(* IEC 61131-3 sources: SRCI_CLIENT_PLC/RobotLibrary/Library/Enumerations/Miscellaneous, 14 files *)

(* ---- AxisUnit.st ---- *)
{attribute 'qualified_only'}
{attribute 'to_string'}
{attribute 'strict'}
// -------------------------------------------------------------------------
//  SRCI Robot Library
// -------------------------------------------------------------------------
//
//  Object:      AxisUnit
//  Author:      Thorsten Brach
//  Date:        2025-03-23
//
//  Description:
//
//
//  Copyright:
//    (C) 2025 Thorsten Brach. All rights reserved
//             Licensed under the MIT License.
//
//  Disclaimer:
//    This project is provided without any guarantee and can be used for
//    private and commercial purposes. Any use is at the user’s
//    own risk and responsibility.
//
// -------------------------------------------------------------------------
TYPE AxisUnit :
(
  /// Axis unit is in degree [°]
	DEG := 0,
  /// Axis unit is in milli meter [mm]
	MM  := 1
)USINT;
END_TYPE

(* ---- CircPlane.st ---- *)
{attribute 'qualified_only'}
{attribute 'to_string'}
{attribute 'strict'}
// -------------------------------------------------------------------------
//  SRCI Robot Library
// -------------------------------------------------------------------------
//
//  Object:      CircPlane
//  Author:      Thorsten Brach
//  Date:        2024-06-01
//
//  Description:
//
//
//  Copyright:
//    (C) 2024 Thorsten Brach. All rights reserved
//             Licensed under the MIT License.
//
//  Disclaimer:
//    This project is provided without any guarantee and can be used for
//    private and commercial purposes. Any use is at the user’s
//    own risk and responsibility.
//
// -------------------------------------------------------------------------
TYPE CircPlane :
(
  /// x-z-plane
  XZ_PLANE := 0,
  /// y-z-plane
  YZ_PLANE := 1,
  /// x-y-plane
  XY_PLANE := 2
)SINT;
END_TYPE

(* ---- ComDirection.st ---- *)
{attribute 'qualified_only'}
{attribute 'to_string'}
{attribute 'strict'}
// -------------------------------------------------------------------------
//  SRCI Robot Library
// -------------------------------------------------------------------------
//
//  Object:      ComDirection
//  Author:      Thorsten Brach
//  Date:        2025-03-23
//
//  Description:
//
//
//  Copyright:
//    (C) 2025 Thorsten Brach. All rights reserved
//             Licensed under the MIT License.
//
//  Disclaimer:
//    This project is provided without any guarantee and can be used for
//    private and commercial purposes. Any use is at the user’s
//    own risk and responsibility.
//
// -------------------------------------------------------------------------
TYPE ComDirection :
(
  // communication direction PLC to Robot
	PLC_TO_ROB := 0,
  // communication direction Robot to PLC
	ROB_TO_PLC := 1
);
END_TYPE

(* ---- ControlHalfByte.st ---- *)
{attribute 'qualified_only'}
{attribute 'to_string'}
// -------------------------------------------------------------------------
//  SRCI Robot Library
// -------------------------------------------------------------------------
//
//  Object:      ControlHalfByte
//  Author:      Thorsten Brach
//  Date:        2024-06-01
//
//  Description:
//
//
//  Copyright:
//    (C) 2024 Thorsten Brach. All rights reserved
//             Licensed under the MIT License.
//
//  Disclaimer:
//    This project is provided without any guarantee and can be used for
//    private and commercial purposes. Any use is at the user’s
//    own risk and responsibility.
//
// -------------------------------------------------------------------------
TYPE ControlHalfByte :
(
  /// Default value, no control active
  NONE := 0,
  /// Initialization is requested by the client
  INITIALIZE := 1,
  /// Resume of operation is requested by the client
  RESUME := 2,
  /// Resetting of the RC is requested by the client. The RC must stop the motion, and clear all state.
  RESET := 3,
  /// Acknowledgement of a telegram state error
  ACK_ERROR := 4,
  /// Signaling that a client error occurred. The Server must respond by setting its RI state to NOT_INITIALIZED
  CLIENT_ERROR := 5
)BYTE;
END_TYPE

(* ---- ErrorReaction.st ---- *)
{attribute 'qualified_only'}
{attribute 'to_string'}
// -------------------------------------------------------------------------
//  SRCI Robot Library
// -------------------------------------------------------------------------
//
//  Object:      ErrorReaction
//  Author:      Thorsten Brach
//  Date:        2024-06-01
//
//  Description:
//
//
//  Copyright:
//    (C) 2024 Thorsten Brach. All rights reserved
//             Licensed under the MIT License.
//
//  Disclaimer:
//    This project is provided without any guarantee and can be used for
//    private and commercial purposes. Any use is at the user’s
//    own risk and responsibility.
//
// -------------------------------------------------------------------------
TYPE ErrorReaction :
(
  /// Abort and move Abort active move command and delete commands buffered in sequence Move robot by specified ErrorVector
  ABORT_AND_MOVE := 0,
  /// 1: Abort
  /// Abort active move command and delete commands buffered in sequence
  /// No additional movements
  ABORT := 1,
  /// 2: No reaction
  /// Error event is ignored by active move command
  NO_REACTION := 2
)USINT;
END_TYPE

(* ---- LoadMeasurementSteps.st ---- *)
{attribute 'qualified_only'}
{attribute 'to_string'}
// -------------------------------------------------------------------------
//  SRCI Robot Library
// -------------------------------------------------------------------------
//
//  Object:      LoadMeasurementSteps
//  Author:      Thorsten Brach
//  Date:        2024-06-01
//
//  Description:
//
//
//  Copyright:
//    (C) 2024 Thorsten Brach. All rights reserved
//             Licensed under the MIT License.
//
//  Disclaimer:
//    This project is provided without any guarantee and can be used for
//    private and commercial purposes. Any use is at the user’s
//    own risk and responsibility.
//
// -------------------------------------------------------------------------
TYPE LoadMeasurementSteps :
(
  /// • 0: Reset (default)
  /// Delete all positions saved on the RC
  RESET := 0,
  /// • 1: First position
  /// Save the first position for the load estimation with the required data
  FIRST_POSITION := 1,
  /// • 2: Second position
  /// Save the second position for the load estimation with the required data
  SECOND_POSITION := 2,
  /// • 3: Third position
  /// Save the third position for the load estimation with the required data
  THIRD_POSITION := 3,
  /// • 4: Fourth position
  /// Save the fourth position for the load estimation with the required data
  FOURTH_POSITION := 4,
  /// • 99: Load calculation
  /// Start the load calculation with the data saved in the four positions
  LOAD_CALCULATION := 99
)USINT;
END_TYPE

(* ---- PathChoice.st ---- *)
{attribute 'qualified_only'}
{attribute 'to_string'}
// -------------------------------------------------------------------------
//  SRCI Robot Library
// -------------------------------------------------------------------------
//
//  Object:      PathChoice
//  Author:      Thorsten Brach
//  Date:        2024-06-01
//
//  Description:
//
//
//  Copyright:
//    (C) 2024 Thorsten Brach. All rights reserved
//             Licensed under the MIT License.
//
//  Disclaimer:
//    This project is provided without any guarantee and can be used for
//    private and commercial purposes. Any use is at the user’s
//    own risk and responsibility.
//
// -------------------------------------------------------------------------
TYPE PathChoice :
(
  /// Clockwise movement of the circular path
  CLOCKWISE := 0,
  /// Counterclockwise movement of the circular path
  COUNTERCLOCKWISE := 1
)BYTE;
END_TYPE

(* ---- ReferenceElement.st ---- *)
{attribute 'qualified_only'}
{attribute 'to_string'}
// -------------------------------------------------------------------------
//  SRCI Robot Library
// -------------------------------------------------------------------------
//
//  Object:      ReferenceElement
//  Author:      Thorsten Brach
//  Date:        2024-06-01
//
//  Description:
//
//
//  Copyright:
//    (C) 2024 Thorsten Brach. All rights reserved
//             Licensed under the MIT License.
//
//  Disclaimer:
//    This project is provided without any guarantee and can be used for
//    private and commercial purposes. Any use is at the user’s
//    own risk and responsibility.
//
// -------------------------------------------------------------------------
TYPE ReferenceElement :
(
  /// 0 (default): Not used
  NOT_USED := 0,
  /// 1: X-Axis
  X_AXIS := 1,
  /// 2: Y-Axis
  Y_AXIS := 2,
  /// 3: Z-Axis
  Z_AXIS := 3,
  /// 4: XY-Plane
  XY_PLANE := 4,
  /// 5: XZ-Plane
  XZ_PLANE := 5,
  /// 6: YZ-Plane
  YZ_PLANE := 6
)USINT;
END_TYPE

(* ---- Severity.st ---- *)
{attribute 'qualified_only'}
{attribute 'to_string'}
// -------------------------------------------------------------------------
//  SRCI Robot Library
// -------------------------------------------------------------------------
//
//  Object:      Severity
//  Author:      Thorsten Brach
//  Date:        2024-06-01
//
//  Description:
//
//
//  Copyright:
//    (C) 2024 Thorsten Brach. All rights reserved
//             Licensed under the MIT License.
//
//  Disclaimer:
//    This project is provided without any guarantee and can be used for
//    private and commercial purposes. Any use is at the user’s
//    own risk and responsibility.
//
// -------------------------------------------------------------------------
TYPE Severity :
(
  /// No events will be logged
  DEACTIVATE  := 0,
  /// Debug message
  /// • No user action required
  DEBUG := 4,
  /// Informative message
  /// • No user action required
  INFO := 5,
  /// Warning message
  /// • User action will be required at some point
  WARNING := 20,
  /// Error message
  /// • User action required immediately
  ERROR := 28,
  ///  Fatal error message
  /// • User action required immediately
  /// • Reinitialization OF RI required
  FATAL_ERROR := 29
)SINT;
END_TYPE

(* ---- SyncDirection.st ---- *)
{attribute 'qualified_only'}
{attribute 'to_string'}
// -------------------------------------------------------------------------
//  SRCI Robot Library
// -------------------------------------------------------------------------
//
//  Object:      SyncDirection
//  Author:      Thorsten Brach
//  Date:        2024-06-01
//
//  Description:
//
//
//  Copyright:
//    (C) 2024 Thorsten Brach. All rights reserved
//             Licensed under the MIT License.
//
//  Disclaimer:
//    This project is provided without any guarantee and can be used for
//    private and commercial purposes. Any use is at the user’s
//    own risk and responsibility.
//
// -------------------------------------------------------------------------
TYPE SyncDirection :
(
  /// No synchronization will be executed
  NO_SYNC := 0,
  /// Server data will be overwritten immediately by client data
  PLC_TO_ROB := 1,
  /// Client data will be overwritten immediately by server data
  ROB_TO_PLC := 2,
  /// Server or client data will be overwritten immediately by changed data
  AUTOMATIC := 3
);
END_TYPE

(* ---- SyncReaction.st ---- *)
{attribute 'qualified_only'}
{attribute 'to_string'}
// -------------------------------------------------------------------------
//  SRCI Robot Library
// -------------------------------------------------------------------------
//
//  Object:      SyncReaction
//  Author:      Thorsten Brach
//  Date:        2024-06-01
//
//  Description:
//
//
//  Copyright:
//    (C) 2024 Thorsten Brach. All rights reserved
//             Licensed under the MIT License.
//
//  Disclaimer:
//    This project is provided without any guarantee and can be used for
//    private and commercial purposes. Any use is at the user’s
//    own risk and responsibility.
//
// -------------------------------------------------------------------------
TYPE SyncReaction :
(
  /// • System behavior unaffected
  NO_REACTION := 0,
  /// • No automatic disable
  /// • Reaction will only apply when RA is disabled
  /// • RA can only be enabled if client and server are synchronized
  NO_AUTOMATIC_DISABLE := 1,
  /// • No automatic disable
  /// • RA can only be enabled if client and server are synchronized
  /// • RA sequence state will change to interrupted when no command is buffered in the active sequence
  /// • Continuation is only possible if client and server are synchronized
  INTERRUPT_WHEN_SEQUENCE_IS_EMPTY := 2,
  /// • No automatic disable
  /// • RA can only be enabled if client and server are synchronized
  /// • RA sequence state will change to interrupted
  /// • Continuation is only possible if client and server are synchronized
  IMMEDIATE_INTERRUPT := 3
)USINT;
END_TYPE

(* ---- SyncTime.st ---- *)
{attribute 'qualified_only'}
{attribute 'to_string'}
// -------------------------------------------------------------------------
//  SRCI Robot Library
// -------------------------------------------------------------------------
//
//  Object:      SyncTime
//  Author:      Thorsten Brach
//  Date:        2025-04-13
//
//  Description:
//
//
//  Copyright:
//    (C) 2025 Thorsten Brach. All rights reserved
//             Licensed under the MIT License.
//
//  Disclaimer:
//    This project is provided without any guarantee and can be used for
//    private and commercial purposes. Any use is at the user’s
//    own risk and responsibility.
//
// -------------------------------------------------------------------------
TYPE SyncTime :
(
  /// Synchronization during startup
	DURING_START_UP := 0,
  /// Synchronization after startup
  AFTER_START_UP := 1
)DINT;
END_TYPE

(* ---- TriggerCondition.st ---- *)
{attribute 'qualified_only'}
{attribute 'to_string'}
// -------------------------------------------------------------------------
//  SRCI Robot Library
// -------------------------------------------------------------------------
//
//  Object:      TriggerCondition
//  Author:      Thorsten Brach
//  Date:        2024-06-01
//
//  Description:
//
//
//  Copyright:
//    (C) 2024 Thorsten Brach. All rights reserved
//             Licensed under the MIT License.
//
//  Disclaimer:
//    This project is provided without any guarantee and can be used for
//    private and commercial purposes. Any use is at the user’s
//    own risk and responsibility.
//
// -------------------------------------------------------------------------
TYPE TriggerCondition :
(
  /// 5: Time in ms  - point reference is target position
  TARGET_POSITION_TIME_MS := -5,
  /// 4: TCP velocity in mm/s - point reference is target position
  TARGET_POSITION_TCP_VELOCITY_ABSOLUTE := -4,
  /// 3: TCP velocity in % of reference velocity - point reference is target position
  TARGET_POSITION_TCP_VELOCITY_PERCENT := -3,
  /// 2: Distance in mm of trajectory - point reference is target position
  TARGET_POSITION_DISTANCE_ABSOLUTE := -2,
  /// 1: Distance in % of trajectory - point reference is target position
  TARGET_POSITION_DISTANCE_PERCENT := -1,
  /// 0: Undfined
  UNDEFINED := 0,
  /// 1: Distance in % of trajectory - point reference is start position
  START_POSITION_DISTANCE_PERCENT := 1,
  /// 2: Distance in mm of trajectory - point reference is start position
  START_POSITION_DISTANCE_ABSOLUTE := 2,
  /// 3: TCP velocity in % of reference velocity - point reference is start position
  START_POSITION_TCP_VELOCITY_PERCENT := 3,
  /// 4: TCP velocity in mm/s - point reference is start position
  START_POSITION_TCP_VELOCITY_ABSOLUTE := 4, // ST-FIX F174: typo in the element name (spec 6.5.17: '4: TCP velocity in mm/s')
  /// 5: Time in ms - point reference is start position
  START_POSITION_TIME_MS := 5
)SINT;
END_TYPE

(* ---- UnitLimitAxis.st ---- *)
{attribute 'qualified_only'}
{attribute 'to_string'}
// -------------------------------------------------------------------------
//  SRCI Robot Library
// -------------------------------------------------------------------------
//
//  Object:      UnitLimitAxis
//  Author:      Thorsten Brach
//  Date:        2025-02-23
//
//  Description:
//
//
//  Copyright:
//    (C) 2025 Thorsten Brach. All rights reserved
//             Licensed under the MIT License.
//
//  Disclaimer:
//    This project is provided without any guarantee and can be used for
//    private and commercial purposes. Any use is at the user’s
//    own risk and responsibility.
//
// -------------------------------------------------------------------------

TYPE UnitLimitAxis :
(
  /// Percentage (%) (default)
	PERCENTAGE  := 0,
  /// Newton meter (Nm)
  NEWTONMETER := 1,
  /// Milliampere (mA)
  MILLIAMPERE := 2
)USINT;
END_TYPE
